// Generated by voz_llm_plc_agent
// Target: Siemens TIA Portal V18 - SCL external source
// Review and compile before any download to physical hardware.

FUNCTION_BLOCK "PLC_PRG"
{ S7_Optimized_Access := 'TRUE' }
VERSION : 0.1
VAR_INPUT
   I_Request_Contactor_A : Bool := FALSE;
   I_Request_Contactor_B : Bool := FALSE;
   I_Emergency : Bool := FALSE;
END_VAR
VAR_OUTPUT
   Q_Contactor_A : Bool := FALSE;
   Q_Contactor_B : Bool := FALSE;
END_VAR
BEGIN
(* Enclavamiento mutuo: cada contactor sigue su propia orden y nunca se activan los dos a la vez *)
(* (el contactor que ya esta activo conserva la prioridad mientras su orden siga presente). *)
IF #I_Emergency THEN
    #Q_Contactor_A := FALSE;
    #Q_Contactor_B := FALSE;
ELSE
    #Q_Contactor_A := #I_Request_Contactor_A AND NOT #Q_Contactor_B;
    #Q_Contactor_B := #I_Request_Contactor_B AND NOT #Q_Contactor_A;
END_IF;
(* Invariante de seguridad: #Q_Contactor_A, #Q_Contactor_B nunca activas a la vez *)
IF (#Q_Contactor_A AND #Q_Contactor_B) THEN
    #Q_Contactor_A := FALSE;
    #Q_Contactor_B := FALSE;
END_IF;
END_FUNCTION_BLOCK

DATA_BLOCK "DB_PLC_PRG"
{ S7_Optimized_Access := 'TRUE' }
VERSION : 0.1
NON_RETAIN
"PLC_PRG"
BEGIN
END_DATA_BLOCK

ORGANIZATION_BLOCK "Main"
{ S7_Optimized_Access := 'TRUE' }
VERSION : 0.1
BEGIN
   "DB_PLC_PRG"(
      I_Request_Contactor_A := "I_Request_Contactor_A",
      I_Request_Contactor_B := "I_Request_Contactor_B",
      I_Emergency := "I_Emergency",
      Q_Contactor_A => "Q_Contactor_A",
      Q_Contactor_B => "Q_Contactor_B"
   );
END_ORGANIZATION_BLOCK
